FUNCTION_BLOCK basicUCT (* Logica unica da UCT Fast (Modbus TCP) e da bomba de gordura com a valvula de lavagem *)
  (* Standard: 61499-2 *)
  (* Version 1.7, 04/11/2026, Hidryco, Hidryco, 1.7: stsLigado para a IO List da Nereda. 1.6: nivel da peneira e velocidades da UCT em % direto (0-100); o 0-16000 da tabela e so o limite do registrador. IHM em Hz (60 Hz = 100 %). 1.5: velocidades dos equipamentos da UCT e da bomba de gordura em Hz (16000 = 60 Hz); conversao no CLP. 1.4: CNF_HMI tambem sai quando muda so a palavra de disponibilidade (STS_HABILITADA). 1.0: UCT Fast (memorial PR-809) por Modbus TCP - leitura de estado, comandos manuais e automaticos por evento, reset, disponibilidade para a EEE Bruto, bomba de gordura e valvula de lavagem *)
  PACKAGE Hidryco.HidrycoLib;
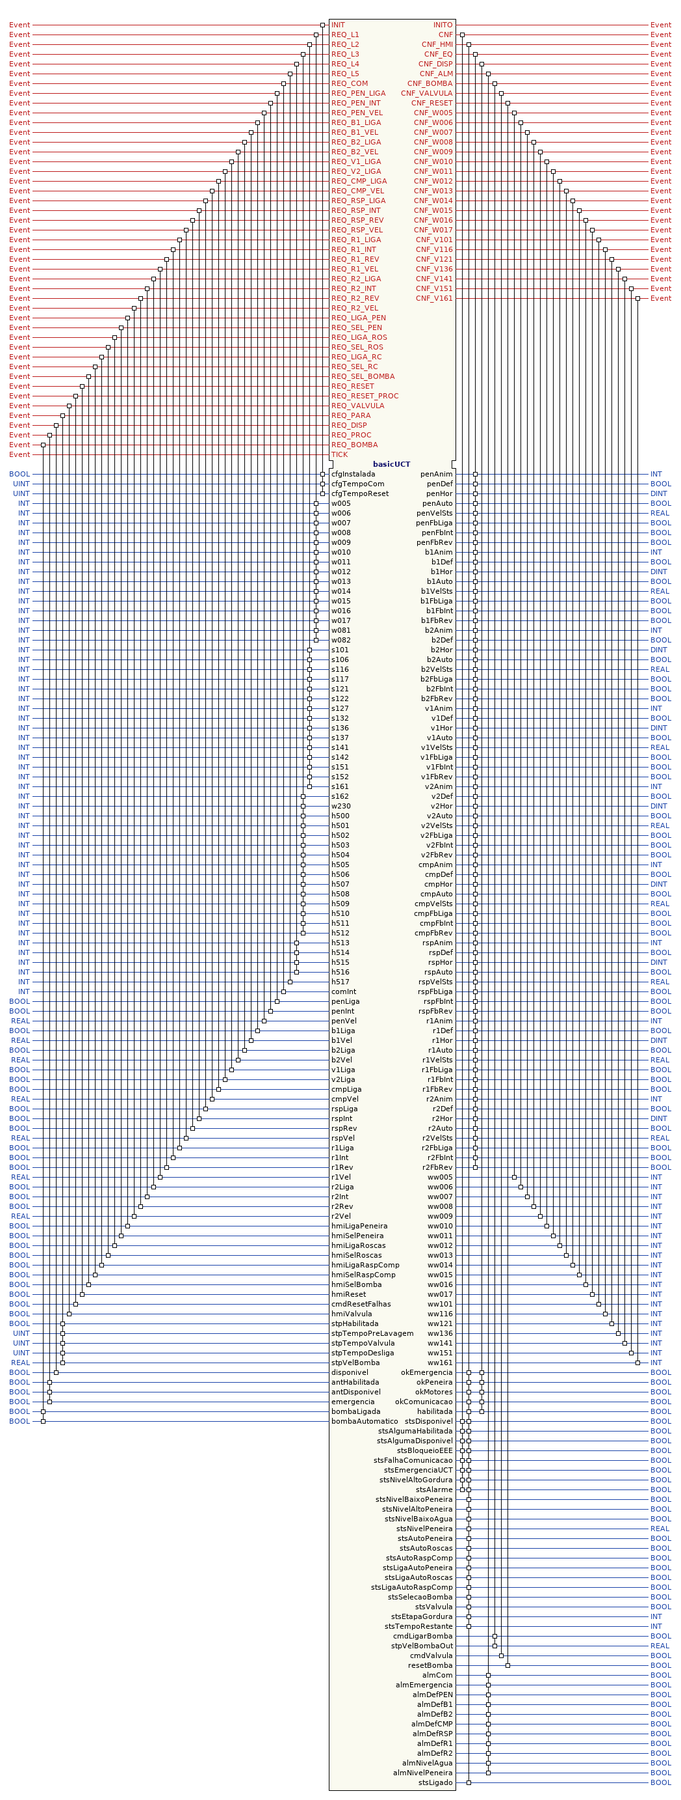
  EVENT_INPUT
    INIT WITH cfgInstalada, cfgTempoCom, cfgTempoReset; (* Inicializacao *)
    REQ_L1 WITH w005, w006, w007, w008, w009, w010, w011, w012, w013, w014, w015, w016, w017, w081, w082; (* Leitura Modbus (grupo 1) *)
    REQ_L2 WITH s101, s106, s116, s117, s121, s122, s127, s132, s136, s137, s141, s142, s151, s152, s161; (* Leitura Modbus (grupo 2) *)
    REQ_L3 WITH s162, w230, h500, h501, h502, h503, h504, h505, h506, h507, h508, h509, h510, h511, h512; (* Leitura Modbus (grupo 3) *)
    REQ_L4 WITH h513, h514, h515, h516; (* Leitura Modbus (grupo 4) *)
    REQ_L5 WITH h517; (* Leitura Modbus (grupo 5) *)
    REQ_COM WITH comInt; (* Comunicacao *)
    REQ_PEN_LIGA WITH penLiga; (* Peneira rotativa: liga manual *)
    REQ_PEN_INT WITH penInt; (* Peneira rotativa: intermitente *)
    REQ_PEN_VEL WITH penVel; (* Peneira rotativa: velocidade (%) *)
    REQ_B1_LIGA WITH b1Liga; (* Bomba 1 de higienização da peneira: liga manual *)
    REQ_B1_VEL WITH b1Vel; (* Bomba 1 de higienização da peneira: velocidade (%) *)
    REQ_B2_LIGA WITH b2Liga; (* Bomba 2 de higienização da peneira: liga manual *)
    REQ_B2_VEL WITH b2Vel; (* Bomba 2 de higienização da peneira: velocidade (%) *)
    REQ_V1_LIGA WITH v1Liga; (* Válvula 1 - higienização do cesto da peneira: liga manual *)
    REQ_V2_LIGA WITH v2Liga; (* Válvula 2 - higienização da rosca da peneira: liga manual *)
    REQ_CMP_LIGA WITH cmpLiga; (* Compressor de ar: liga manual *)
    REQ_CMP_VEL WITH cmpVel; (* Compressor de ar: velocidade (%) *)
    REQ_RSP_LIGA WITH rspLiga; (* Raspador de gordura: liga manual *)
    REQ_RSP_INT WITH rspInt; (* Raspador de gordura: intermitente *)
    REQ_RSP_REV WITH rspRev; (* Raspador de gordura: reversao *)
    REQ_RSP_VEL WITH rspVel; (* Raspador de gordura: velocidade (%) *)
    REQ_R1_LIGA WITH r1Liga; (* Rosca 1 - horizontal: liga manual *)
    REQ_R1_INT WITH r1Int; (* Rosca 1 - horizontal: intermitente *)
    REQ_R1_REV WITH r1Rev; (* Rosca 1 - horizontal: reversao *)
    REQ_R1_VEL WITH r1Vel; (* Rosca 1 - horizontal: velocidade (%) *)
    REQ_R2_LIGA WITH r2Liga; (* Rosca 2 - inclinada: liga manual *)
    REQ_R2_INT WITH r2Int; (* Rosca 2 - inclinada: intermitente *)
    REQ_R2_REV WITH r2Rev; (* Rosca 2 - inclinada: reversao *)
    REQ_R2_VEL WITH r2Vel; (* Rosca 2 - inclinada: velocidade (%) *)
    REQ_LIGA_PEN WITH hmiLigaPeneira; (* cmdLigaSubsistemaPeneira *)
    REQ_SEL_PEN WITH hmiSelPeneira; (* cmdSelecaoSubsistemaPeneira *)
    REQ_LIGA_ROS WITH hmiLigaRoscas; (* cmdLigaSubsistemaRoscas *)
    REQ_SEL_ROS WITH hmiSelRoscas; (* cmdSelecaoSubsistemaRoscas *)
    REQ_LIGA_RC WITH hmiLigaRaspComp; (* cmdLigaSubsistemaRaspComp *)
    REQ_SEL_RC WITH hmiSelRaspComp; (* cmdSelecaoSubsistemaRaspComp *)
    REQ_SEL_BOMBA WITH hmiSelBomba; (* cmdSelecaoBombaHigienizacao *)
    REQ_RESET WITH hmiReset; (* Reset pela IHM *)
    REQ_RESET_PROC WITH cmdResetFalhas; (* Reset pelo processo *)
    REQ_VALVULA WITH hmiValvula; (* Valvula de lavagem manual *)
    REQ_PARA WITH stpHabilitada, stpTempoPreLavagem, stpTempoValvula, stpTempoDesliga, stpVelBomba; (* Parametros (persistentes) *)
    REQ_DISP WITH disponivel; (* Resultado do AND de disponibilidade *)
    REQ_PROC WITH antHabilitada, antDisponivel, emergencia; (* Cadeia das UCTs e emergencia *)
    REQ_BOMBA WITH bombaLigada, bombaAutomatico; (* Estado da bomba de gordura *)
    TICK; (* Base de tempo de 1 s (E_CYCLE) *)
  END_EVENT
  EVENT_OUTPUT
    INITO; (* Inicializacao concluida *)
    CNF WITH stsDisponivel, stsAlgumaHabilitada, stsAlgumaDisponivel, stsBloqueioEEE, stsFalhaComunicacao, stsEmergenciaUCT, stsNivelAltoGordura, stsAlarme; (* Processo (na mudanca) *)
    CNF_HMI WITH stsDisponivel, stsAlgumaHabilitada, stsAlgumaDisponivel, stsBloqueioEEE, stsFalhaComunicacao, stsEmergenciaUCT, stsNivelAltoGordura, stsAlarme, stsNivelBaixoPeneira, stsNivelAltoPeneira, stsNivelBaixoAgua, stsNivelPeneira, stsAutoPeneira, stsAutoRoscas, stsAutoRaspComp, stsLigaAutoPeneira, stsLigaAutoRoscas, stsLigaAutoRaspComp, stsSelecaoBomba, stsValvula, stsEtapaGordura, stsTempoRestante, okEmergencia, okPeneira, okMotores, okComunicacao, habilitada, stsLigado; (* IHM da UCT (na mudanca) *)
    CNF_EQ WITH penAnim, penDef, penHor, penAuto, penVelSts, penFbLiga, penFbInt, penFbRev, b1Anim, b1Def, b1Hor, b1Auto, b1VelSts, b1FbLiga, b1FbInt, b1FbRev, b2Anim, b2Def, b2Hor, b2Auto, b2VelSts, b2FbLiga, b2FbInt, b2FbRev, v1Anim, v1Def, v1Hor, v1Auto, v1VelSts, v1FbLiga, v1FbInt, v1FbRev, v2Anim, v2Def, v2Hor, v2Auto, v2VelSts, v2FbLiga, v2FbInt, v2FbRev, cmpAnim, cmpDef, cmpHor, cmpAuto, cmpVelSts, cmpFbLiga, cmpFbInt, cmpFbRev, rspAnim, rspDef, rspHor, rspAuto, rspVelSts, rspFbLiga, rspFbInt, rspFbRev, r1Anim, r1Def, r1Hor, r1Auto, r1VelSts, r1FbLiga, r1FbInt, r1FbRev, r2Anim, r2Def, r2Hor, r2Auto, r2VelSts, r2FbLiga, r2FbInt, r2FbRev; (* IHM dos equipamentos (na mudanca) *)
    CNF_DISP WITH okEmergencia, okPeneira, okMotores, okComunicacao, habilitada; (* Condicoes para o AND de disponibilidade (na mudanca) *)
    CNF_ALM WITH almCom, almEmergencia, almDefPEN, almDefB1, almDefB2, almDefCMP, almDefRSP, almDefR1, almDefR2, almNivelAgua, almNivelPeneira; (* Alarmes para os ALARM_BIT (na mudanca) *)
    CNF_BOMBA WITH cmdLigarBomba, stpVelBombaOut; (* Bomba de gordura (na mudanca) *)
    CNF_VALVULA WITH cmdValvula; (* Valvula de lavagem (na mudanca) *)
    CNF_RESET WITH resetBomba; (* Reset da bomba de gordura *)
    CNF_W005 WITH ww005; (* Escreve 40005 na UCT *)
    CNF_W006 WITH ww006; (* Escreve 40006 na UCT *)
    CNF_W007 WITH ww007; (* Escreve 40007 na UCT *)
    CNF_W008 WITH ww008; (* Escreve 40008 na UCT *)
    CNF_W009 WITH ww009; (* Escreve 40009 na UCT *)
    CNF_W010 WITH ww010; (* Escreve 40010 na UCT *)
    CNF_W011 WITH ww011; (* Escreve 40011 na UCT *)
    CNF_W012 WITH ww012; (* Escreve 40012 na UCT *)
    CNF_W013 WITH ww013; (* Escreve 40013 na UCT *)
    CNF_W014 WITH ww014; (* Escreve 40014 na UCT *)
    CNF_W015 WITH ww015; (* Escreve 40015 na UCT *)
    CNF_W016 WITH ww016; (* Escreve 40016 na UCT *)
    CNF_W017 WITH ww017; (* Escreve 40017 na UCT *)
    CNF_V101 WITH ww101; (* Escreve 40101 na UCT *)
    CNF_V116 WITH ww116; (* Escreve 40116 na UCT *)
    CNF_V121 WITH ww121; (* Escreve 40121 na UCT *)
    CNF_V136 WITH ww136; (* Escreve 40136 na UCT *)
    CNF_V141 WITH ww141; (* Escreve 40141 na UCT *)
    CNF_V151 WITH ww151; (* Escreve 40151 na UCT *)
    CNF_V161 WITH ww161; (* Escreve 40161 na UCT *)
  END_EVENT
  VAR_INPUT
    cfgInstalada : BOOL := TRUE; (* FALSE = UCT ainda nao existe em campo (sem comunicacao, sem alarmes, fora do bloqueio da EEE) *)
    cfgTempoCom : UINT := 10; (* Tempo (s) sem comunicacao com a UCT para confirmar a falha *)
    cfgTempoReset : UINT := 2; (* Tempo (s) do pulso de reset escrito na UCT (40005.3) *)
    w005 : INT; (* Modbus UCT 40005 *)
    w006 : INT; (* Modbus UCT 40006 *)
    w007 : INT; (* Modbus UCT 40007 *)
    w008 : INT; (* Modbus UCT 40008 *)
    w009 : INT; (* Modbus UCT 40009 *)
    w010 : INT; (* Modbus UCT 40010 *)
    w011 : INT; (* Modbus UCT 40011 *)
    w012 : INT; (* Modbus UCT 40012 *)
    w013 : INT; (* Modbus UCT 40013 *)
    w014 : INT; (* Modbus UCT 40014 *)
    w015 : INT; (* Modbus UCT 40015 *)
    w016 : INT; (* Modbus UCT 40016 *)
    w017 : INT; (* Modbus UCT 40017 *)
    w081 : INT; (* Modbus UCT 40081 *)
    w082 : INT; (* Modbus UCT 40082 *)
    s101 : INT; (* Modbus UCT 40101 *)
    s106 : INT; (* Modbus UCT 40106 *)
    s116 : INT; (* Modbus UCT 40116 *)
    s117 : INT; (* Modbus UCT 40117 *)
    s121 : INT; (* Modbus UCT 40121 *)
    s122 : INT; (* Modbus UCT 40122 *)
    s127 : INT; (* Modbus UCT 40127 *)
    s132 : INT; (* Modbus UCT 40132 *)
    s136 : INT; (* Modbus UCT 40136 *)
    s137 : INT; (* Modbus UCT 40137 *)
    s141 : INT; (* Modbus UCT 40141 *)
    s142 : INT; (* Modbus UCT 40142 *)
    s151 : INT; (* Modbus UCT 40151 *)
    s152 : INT; (* Modbus UCT 40152 *)
    s161 : INT; (* Modbus UCT 40161 *)
    s162 : INT; (* Modbus UCT 40162 *)
    w230 : INT; (* Modbus UCT 40230 *)
    h500 : INT; (* Modbus UCT 40500 *)
    h501 : INT; (* Modbus UCT 40501 *)
    h502 : INT; (* Modbus UCT 40502 *)
    h503 : INT; (* Modbus UCT 40503 *)
    h504 : INT; (* Modbus UCT 40504 *)
    h505 : INT; (* Modbus UCT 40505 *)
    h506 : INT; (* Modbus UCT 40506 *)
    h507 : INT; (* Modbus UCT 40507 *)
    h508 : INT; (* Modbus UCT 40508 *)
    h509 : INT; (* Modbus UCT 40509 *)
    h510 : INT; (* Modbus UCT 40510 *)
    h511 : INT; (* Modbus UCT 40511 *)
    h512 : INT; (* Modbus UCT 40512 *)
    h513 : INT; (* Modbus UCT 40513 *)
    h514 : INT; (* Modbus UCT 40514 *)
    h515 : INT; (* Modbus UCT 40515 *)
    h516 : INT; (* Modbus UCT 40516 *)
    h517 : INT; (* Modbus UCT 40517 *)
    comInt : INT; (* connStatusInt do escravo Modbus da UCT (1 = online) *)
    penLiga : BOOL; (* IHM: Peneira rotativa: liga manual *)
    penInt : BOOL; (* IHM: Peneira rotativa: intermitente *)
    penVel : REAL; (* IHM: Peneira rotativa: velocidade (%) *)
    b1Liga : BOOL; (* IHM: Bomba 1 de higienização da peneira: liga manual *)
    b1Vel : REAL; (* IHM: Bomba 1 de higienização da peneira: velocidade (%) *)
    b2Liga : BOOL; (* IHM: Bomba 2 de higienização da peneira: liga manual *)
    b2Vel : REAL; (* IHM: Bomba 2 de higienização da peneira: velocidade (%) *)
    v1Liga : BOOL; (* IHM: Válvula 1 - higienização do cesto da peneira: liga manual *)
    v2Liga : BOOL; (* IHM: Válvula 2 - higienização da rosca da peneira: liga manual *)
    cmpLiga : BOOL; (* IHM: Compressor de ar: liga manual *)
    cmpVel : REAL; (* IHM: Compressor de ar: velocidade (%) *)
    rspLiga : BOOL; (* IHM: Raspador de gordura: liga manual *)
    rspInt : BOOL; (* IHM: Raspador de gordura: intermitente *)
    rspRev : BOOL; (* IHM: Raspador de gordura: reversao *)
    rspVel : REAL; (* IHM: Raspador de gordura: velocidade (%) *)
    r1Liga : BOOL; (* IHM: Rosca 1 - horizontal: liga manual *)
    r1Int : BOOL; (* IHM: Rosca 1 - horizontal: intermitente *)
    r1Rev : BOOL; (* IHM: Rosca 1 - horizontal: reversao *)
    r1Vel : REAL; (* IHM: Rosca 1 - horizontal: velocidade (%) *)
    r2Liga : BOOL; (* IHM: Rosca 2 - inclinada: liga manual *)
    r2Int : BOOL; (* IHM: Rosca 2 - inclinada: intermitente *)
    r2Rev : BOOL; (* IHM: Rosca 2 - inclinada: reversao *)
    r2Vel : REAL; (* IHM: Rosca 2 - inclinada: velocidade (%) *)
    hmiLigaPeneira : BOOL; (* IHM: cmdLigaSubsistemaPeneira *)
    hmiSelPeneira : BOOL; (* IHM: cmdSelecaoSubsistemaPeneira *)
    hmiLigaRoscas : BOOL; (* IHM: cmdLigaSubsistemaRoscas *)
    hmiSelRoscas : BOOL; (* IHM: cmdSelecaoSubsistemaRoscas *)
    hmiLigaRaspComp : BOOL; (* IHM: cmdLigaSubsistemaRaspComp *)
    hmiSelRaspComp : BOOL; (* IHM: cmdSelecaoSubsistemaRaspComp *)
    hmiSelBomba : BOOL; (* IHM: cmdSelecaoBombaHigienizacao *)
    hmiReset : BOOL; (* IHM: reset (reconhece e reseta a UCT e a bomba de gordura) *)
    cmdResetFalhas : BOOL; (* Processo: reset (com E_RESET_FALHAS) *)
    hmiValvula : BOOL; (* IHM: valvula de lavagem aberta (TRUE) / fechada (FALSE) - so com a bomba de gordura fora do automatico *)
    stpHabilitada : BOOL; (* IHM (persistente): UCT habilitada no bloqueio da EEE Bruto (desabilitada nao conta) *)
    stpTempoPreLavagem : UINT; (* IHM (persistente): Tempo (s) com a valvula de lavagem aberta antes de ligar a bomba de gordura (0 = liga junto) *)
    stpTempoValvula : UINT; (* IHM (persistente): Tempo (s) que a valvula fica aberta depois que a bomba liga (0 = fecha na partida) *)
    stpTempoDesliga : UINT; (* IHM (persistente): Tempo (s) que a bomba de gordura continua ligada depois que o nivel alto do tanque abaixa *)
    stpVelBomba : REAL; (* IHM (persistente): Velocidade da bomba de gordura em automatico (%) *)
    disponivel : BOOL; (* Saida do bloco AND editavel: UCT disponivel *)
    antHabilitada : BOOL; (* UCT anterior na cadeia: alguma UCT habilitada *)
    antDisponivel : BOOL; (* UCT anterior na cadeia: alguma UCT disponivel *)
    emergencia : BOOL; (* Emergencia pelo processo (fecha a valvula de lavagem) *)
    bombaLigada : BOOL; (* Bomba de gordura ligada (Motor_Generico.stsLigado) *)
    bombaAutomatico : BOOL; (* Bomba de gordura em automatico (Motor_Generico.stsAutomatico) *)
  END_VAR
  VAR_OUTPUT
    penAnim : INT; (* Peneira rotativa: 0 desligado, 1 ligado, 2 falha, 3 manutencao, 4 sem comunicacao *)
    penDef : BOOL; (* Peneira rotativa: defeito *)
    penHor : DINT; (* Peneira rotativa: horimetro (h) *)
    penAuto : BOOL; (* Peneira rotativa: subsistema em automatico *)
    penVelSts : REAL; (* Peneira rotativa: velocidade (%) *)
    penFbLiga : BOOL; (* Peneira rotativa: liga em vigor *)
    penFbInt : BOOL; (* Peneira rotativa: intermitente em vigor *)
    penFbRev : BOOL; (* Peneira rotativa: reversao em vigor *)
    b1Anim : INT; (* Bomba 1 de higienização da peneira: 0 desligado, 1 ligado, 2 falha, 3 manutencao, 4 sem comunicacao *)
    b1Def : BOOL; (* Bomba 1 de higienização da peneira: defeito *)
    b1Hor : DINT; (* Bomba 1 de higienização da peneira: horimetro (h) *)
    b1Auto : BOOL; (* Bomba 1 de higienização da peneira: subsistema em automatico *)
    b1VelSts : REAL; (* Bomba 1 de higienização da peneira: velocidade (%) *)
    b1FbLiga : BOOL; (* Bomba 1 de higienização da peneira: liga em vigor *)
    b1FbInt : BOOL; (* Bomba 1 de higienização da peneira: intermitente em vigor *)
    b1FbRev : BOOL; (* Bomba 1 de higienização da peneira: reversao em vigor *)
    b2Anim : INT; (* Bomba 2 de higienização da peneira: 0 desligado, 1 ligado, 2 falha, 3 manutencao, 4 sem comunicacao *)
    b2Def : BOOL; (* Bomba 2 de higienização da peneira: defeito *)
    b2Hor : DINT; (* Bomba 2 de higienização da peneira: horimetro (h) *)
    b2Auto : BOOL; (* Bomba 2 de higienização da peneira: subsistema em automatico *)
    b2VelSts : REAL; (* Bomba 2 de higienização da peneira: velocidade (%) *)
    b2FbLiga : BOOL; (* Bomba 2 de higienização da peneira: liga em vigor *)
    b2FbInt : BOOL; (* Bomba 2 de higienização da peneira: intermitente em vigor *)
    b2FbRev : BOOL; (* Bomba 2 de higienização da peneira: reversao em vigor *)
    v1Anim : INT; (* Válvula 1 - higienização do cesto da peneira: 0 desligado, 1 ligado, 2 falha, 3 manutencao, 4 sem comunicacao *)
    v1Def : BOOL; (* Válvula 1 - higienização do cesto da peneira: defeito *)
    v1Hor : DINT; (* Válvula 1 - higienização do cesto da peneira: horimetro (h) *)
    v1Auto : BOOL; (* Válvula 1 - higienização do cesto da peneira: subsistema em automatico *)
    v1VelSts : REAL; (* Válvula 1 - higienização do cesto da peneira: velocidade (%) *)
    v1FbLiga : BOOL; (* Válvula 1 - higienização do cesto da peneira: liga em vigor *)
    v1FbInt : BOOL; (* Válvula 1 - higienização do cesto da peneira: intermitente em vigor *)
    v1FbRev : BOOL; (* Válvula 1 - higienização do cesto da peneira: reversao em vigor *)
    v2Anim : INT; (* Válvula 2 - higienização da rosca da peneira: 0 desligado, 1 ligado, 2 falha, 3 manutencao, 4 sem comunicacao *)
    v2Def : BOOL; (* Válvula 2 - higienização da rosca da peneira: defeito *)
    v2Hor : DINT; (* Válvula 2 - higienização da rosca da peneira: horimetro (h) *)
    v2Auto : BOOL; (* Válvula 2 - higienização da rosca da peneira: subsistema em automatico *)
    v2VelSts : REAL; (* Válvula 2 - higienização da rosca da peneira: velocidade (%) *)
    v2FbLiga : BOOL; (* Válvula 2 - higienização da rosca da peneira: liga em vigor *)
    v2FbInt : BOOL; (* Válvula 2 - higienização da rosca da peneira: intermitente em vigor *)
    v2FbRev : BOOL; (* Válvula 2 - higienização da rosca da peneira: reversao em vigor *)
    cmpAnim : INT; (* Compressor de ar: 0 desligado, 1 ligado, 2 falha, 3 manutencao, 4 sem comunicacao *)
    cmpDef : BOOL; (* Compressor de ar: defeito *)
    cmpHor : DINT; (* Compressor de ar: horimetro (h) *)
    cmpAuto : BOOL; (* Compressor de ar: subsistema em automatico *)
    cmpVelSts : REAL; (* Compressor de ar: velocidade (%) *)
    cmpFbLiga : BOOL; (* Compressor de ar: liga em vigor *)
    cmpFbInt : BOOL; (* Compressor de ar: intermitente em vigor *)
    cmpFbRev : BOOL; (* Compressor de ar: reversao em vigor *)
    rspAnim : INT; (* Raspador de gordura: 0 desligado, 1 ligado, 2 falha, 3 manutencao, 4 sem comunicacao *)
    rspDef : BOOL; (* Raspador de gordura: defeito *)
    rspHor : DINT; (* Raspador de gordura: horimetro (h) *)
    rspAuto : BOOL; (* Raspador de gordura: subsistema em automatico *)
    rspVelSts : REAL; (* Raspador de gordura: velocidade (%) *)
    rspFbLiga : BOOL; (* Raspador de gordura: liga em vigor *)
    rspFbInt : BOOL; (* Raspador de gordura: intermitente em vigor *)
    rspFbRev : BOOL; (* Raspador de gordura: reversao em vigor *)
    r1Anim : INT; (* Rosca 1 - horizontal: 0 desligado, 1 ligado, 2 falha, 3 manutencao, 4 sem comunicacao *)
    r1Def : BOOL; (* Rosca 1 - horizontal: defeito *)
    r1Hor : DINT; (* Rosca 1 - horizontal: horimetro (h) *)
    r1Auto : BOOL; (* Rosca 1 - horizontal: subsistema em automatico *)
    r1VelSts : REAL; (* Rosca 1 - horizontal: velocidade (%) *)
    r1FbLiga : BOOL; (* Rosca 1 - horizontal: liga em vigor *)
    r1FbInt : BOOL; (* Rosca 1 - horizontal: intermitente em vigor *)
    r1FbRev : BOOL; (* Rosca 1 - horizontal: reversao em vigor *)
    r2Anim : INT; (* Rosca 2 - inclinada: 0 desligado, 1 ligado, 2 falha, 3 manutencao, 4 sem comunicacao *)
    r2Def : BOOL; (* Rosca 2 - inclinada: defeito *)
    r2Hor : DINT; (* Rosca 2 - inclinada: horimetro (h) *)
    r2Auto : BOOL; (* Rosca 2 - inclinada: subsistema em automatico *)
    r2VelSts : REAL; (* Rosca 2 - inclinada: velocidade (%) *)
    r2FbLiga : BOOL; (* Rosca 2 - inclinada: liga em vigor *)
    r2FbInt : BOOL; (* Rosca 2 - inclinada: intermitente em vigor *)
    r2FbRev : BOOL; (* Rosca 2 - inclinada: reversao em vigor *)
    ww005 : INT; (* Palavra escrita na UCT: 40005 *)
    ww006 : INT; (* Palavra escrita na UCT: 40006 *)
    ww007 : INT; (* Palavra escrita na UCT: 40007 *)
    ww008 : INT; (* Palavra escrita na UCT: 40008 *)
    ww009 : INT; (* Palavra escrita na UCT: 40009 *)
    ww010 : INT; (* Palavra escrita na UCT: 40010 *)
    ww011 : INT; (* Palavra escrita na UCT: 40011 *)
    ww012 : INT; (* Palavra escrita na UCT: 40012 *)
    ww013 : INT; (* Palavra escrita na UCT: 40013 *)
    ww014 : INT; (* Palavra escrita na UCT: 40014 *)
    ww015 : INT; (* Palavra escrita na UCT: 40015 *)
    ww016 : INT; (* Palavra escrita na UCT: 40016 *)
    ww017 : INT; (* Palavra escrita na UCT: 40017 *)
    ww101 : INT; (* Palavra escrita na UCT: 40101 *)
    ww116 : INT; (* Palavra escrita na UCT: 40116 *)
    ww121 : INT; (* Palavra escrita na UCT: 40121 *)
    ww136 : INT; (* Palavra escrita na UCT: 40136 *)
    ww141 : INT; (* Palavra escrita na UCT: 40141 *)
    ww151 : INT; (* Palavra escrita na UCT: 40151 *)
    ww161 : INT; (* Palavra escrita na UCT: 40161 *)
    okEmergencia : BOOL; (* UCT sem emergencia *)
    okPeneira : BOOL; (* Peneira sem defeito *)
    okMotores : BOOL; (* Bombas de higienizacao, roscas, raspador e compressor sem defeito *)
    okComunicacao : BOOL; (* Comunicacao com a UCT ok *)
    habilitada : BOOL; (* UCT instalada e habilitada *)
    stsDisponivel : BOOL; (* UCT disponivel (saida do AND) *)
    stsAlgumaHabilitada : BOOL; (* Esta UCT ou alguma anterior habilitada *)
    stsAlgumaDisponivel : BOOL; (* Esta UCT ou alguma anterior disponivel *)
    stsBloqueioEEE : BOOL; (* Bloqueio do automatico da EEE Bruto: ha UCT habilitada e nenhuma disponivel *)
    stsFalhaComunicacao : BOOL; (* Falha de comunicacao com a UCT *)
    stsEmergenciaUCT : BOOL; (* Emergencia acionada na UCT *)
    stsNivelAltoGordura : BOOL; (* Nivel alto do tanque de gordura (UCT) *)
    stsAlarme : BOOL; (* Algum alarme da UCT *)
    stsNivelBaixoPeneira : BOOL; (* Nivel baixo da peneira *)
    stsNivelAltoPeneira : BOOL; (* Nivel alto da peneira *)
    stsNivelBaixoAgua : BOOL; (* Nivel baixo do tanque de agua *)
    stsNivelPeneira : REAL; (* Nivel da peneira (%) *)
    stsAutoPeneira : BOOL; (* Subsistema peneira e higienização em automatico *)
    stsAutoRoscas : BOOL; (* Subsistema roscas em automatico *)
    stsAutoRaspComp : BOOL; (* Subsistema raspador e compressor em automatico *)
    stsLigaAutoPeneira : BOOL; (* Subsistema peneira e higienização: liga automatico em vigor *)
    stsLigaAutoRoscas : BOOL; (* Subsistema roscas: liga automatico em vigor *)
    stsLigaAutoRaspComp : BOOL; (* Subsistema raspador e compressor: liga automatico em vigor *)
    stsSelecaoBomba : BOOL; (* Bomba de higienizacao selecionada: FALSE = bomba 1, TRUE = bomba 2 *)
    stsValvula : BOOL; (* Valvula de lavagem do tanque de gordura aberta *)
    stsEtapaGordura : INT; (* Bomba de gordura: 0 parada, 1 pre-lavagem, 2 bombeando, 3 nivel normal - contando para desligar, 4 fora do automatico *)
    stsTempoRestante : INT; (* Tempo restante (s) da etapa da bomba de gordura *)
    cmdLigarBomba : BOOL; (* Bomba de gordura: liga em automatico (Motor_Generico.cmdLigarAutomatico) *)
    stpVelBombaOut : REAL; (* Bomba de gordura: velocidade em automatico (%) *)
    cmdValvula : BOOL; (* Valvula de lavagem: saida digital (symlink ${PATH}cmdValvulaLavagem) *)
    resetBomba : BOOL; (* Reset da bomba de gordura (com CNF_RESET) *)
    almCom : BOOL; (* ALARM_BIT Falha de comunicação com a UCT *)
    almEmergencia : BOOL; (* ALARM_BIT Emergência acionada na UCT *)
    almDefPEN : BOOL; (* ALARM_BIT Defeito: Peneira rotativa *)
    almDefB1 : BOOL; (* ALARM_BIT Defeito: Bomba 1 de higienização da peneira *)
    almDefB2 : BOOL; (* ALARM_BIT Defeito: Bomba 2 de higienização da peneira *)
    almDefCMP : BOOL; (* ALARM_BIT Defeito: Compressor de ar *)
    almDefRSP : BOOL; (* ALARM_BIT Defeito: Raspador de gordura *)
    almDefR1 : BOOL; (* ALARM_BIT Defeito: Rosca 1 - horizontal *)
    almDefR2 : BOOL; (* ALARM_BIT Defeito: Rosca 2 - inclinada *)
    almNivelAgua : BOOL; (* ALARM_BIT Nível baixo do tanque de água de higienização da UCT *)
    almNivelPeneira : BOOL; (* ALARM_BIT Nível alto na peneira da UCT *)
    stsLigado : BOOL; (* Algum subsistema com liga-automatico (peneira, roscas ou raspador/compressor) *)
  END_VAR
  VAR
    initDone : BOOL;
    initPass : BOOL;
    bComRecebida : BOOL; (* Ja houve leitura do connStatusInt *)
    bLeitura : BOOL; (* Ja houve leitura das palavras de comando *)
    bComOK : BOOL; (* Comunicando agora *)
    uSegCom : UDINT;
    uSegReset : UINT; (* Segundos do pulso de reset *)
    bReset : BOOL;
    w81 : WORD;
    w82 : WORD;
    bNivelAltoG : BOOL; (* Nivel alto do tanque de gordura valido *)
    uEtapa : INT; (* Etapa da bomba de gordura *)
    uSegEtapa : UDINT; (* Segundos na etapa *)
    uSegValv : UDINT; (* Segundos com a bomba ligada *)
    bValvAuto : BOOL; (* Valvula pedida pela sequencia *)
    bMudou : BOOL;
    wD : WORD;
    oldD : WORD := 16#FFFF;
    wP : DWORD;
    oldP : DWORD := 16#FFFFFFFF;
    wA : WORD;
    oldA : WORD := 16#FFFF;
    oldLigB : BOOL;
    oldVelB : REAL := -1.0;
    oldValv : BOOL;
    img005 : WORD; (* Imagem da palavra 40005 (lida da UCT, alterada so no bit comandado) *)
    img006 : WORD; (* Imagem da palavra 40006 (lida da UCT, alterada so no bit comandado) *)
    img007 : WORD; (* Imagem da palavra 40007 (lida da UCT, alterada so no bit comandado) *)
    img008 : WORD; (* Imagem da palavra 40008 (lida da UCT, alterada so no bit comandado) *)
    img009 : WORD; (* Imagem da palavra 40009 (lida da UCT, alterada so no bit comandado) *)
    img010 : WORD; (* Imagem da palavra 40010 (lida da UCT, alterada so no bit comandado) *)
    img011 : WORD; (* Imagem da palavra 40011 (lida da UCT, alterada so no bit comandado) *)
    img012 : WORD; (* Imagem da palavra 40012 (lida da UCT, alterada so no bit comandado) *)
    img013 : WORD; (* Imagem da palavra 40013 (lida da UCT, alterada so no bit comandado) *)
    img014 : WORD; (* Imagem da palavra 40014 (lida da UCT, alterada so no bit comandado) *)
    img015 : WORD; (* Imagem da palavra 40015 (lida da UCT, alterada so no bit comandado) *)
    img016 : WORD; (* Imagem da palavra 40016 (lida da UCT, alterada so no bit comandado) *)
    img017 : WORD; (* Imagem da palavra 40017 (lida da UCT, alterada so no bit comandado) *)
    o_stsNivelPeneira : REAL := -1.0;
    o_stsEtapaGordura : INT := -1;
    o_stsTempoRestante : INT := -1;
    o_penAnim : INT := -1;
    o_penHor : DINT := -1;
    o_penVelSts : REAL := -1.0;
    o_b1Anim : INT := -1;
    o_b1Hor : DINT := -1;
    o_b1VelSts : REAL := -1.0;
    o_b2Anim : INT := -1;
    o_b2Hor : DINT := -1;
    o_b2VelSts : REAL := -1.0;
    o_v1Anim : INT := -1;
    o_v1Hor : DINT := -1;
    o_v1VelSts : REAL := -1.0;
    o_v2Anim : INT := -1;
    o_v2Hor : DINT := -1;
    o_v2VelSts : REAL := -1.0;
    o_cmpAnim : INT := -1;
    o_cmpHor : DINT := -1;
    o_cmpVelSts : REAL := -1.0;
    o_rspAnim : INT := -1;
    o_rspHor : DINT := -1;
    o_rspVelSts : REAL := -1.0;
    o_r1Anim : INT := -1;
    o_r1Hor : DINT := -1;
    o_r1VelSts : REAL := -1.0;
    o_r2Anim : INT := -1;
    o_r2Hor : DINT := -1;
    o_r2VelSts : REAL := -1.0;
    o_penDef : BOOL;
    o_penAuto : BOOL;
    o_penFbLiga : BOOL;
    o_penFbInt : BOOL;
    o_penFbRev : BOOL;
    o_b1Def : BOOL;
    o_b1Auto : BOOL;
    o_b1FbLiga : BOOL;
    o_b1FbInt : BOOL;
    o_b1FbRev : BOOL;
    o_b2Def : BOOL;
    o_b2Auto : BOOL;
    o_b2FbLiga : BOOL;
    o_b2FbInt : BOOL;
    o_b2FbRev : BOOL;
    o_v1Def : BOOL;
    o_v1Auto : BOOL;
    o_v1FbLiga : BOOL;
    o_v1FbInt : BOOL;
    o_v1FbRev : BOOL;
    o_v2Def : BOOL;
    o_v2Auto : BOOL;
    o_v2FbLiga : BOOL;
    o_v2FbInt : BOOL;
    o_v2FbRev : BOOL;
    o_cmpDef : BOOL;
    o_cmpAuto : BOOL;
    o_cmpFbLiga : BOOL;
    o_cmpFbInt : BOOL;
    o_cmpFbRev : BOOL;
    o_rspDef : BOOL;
    o_rspAuto : BOOL;
    o_rspFbLiga : BOOL;
    o_rspFbInt : BOOL;
    o_rspFbRev : BOOL;
    o_r1Def : BOOL;
    o_r1Auto : BOOL;
    o_r1FbLiga : BOOL;
    o_r1FbInt : BOOL;
    o_r1FbRev : BOOL;
    o_r2Def : BOOL;
    o_r2Auto : BOOL;
    o_r2FbLiga : BOOL;
    o_r2FbInt : BOOL;
    o_r2FbRev : BOOL;
  END_VAR
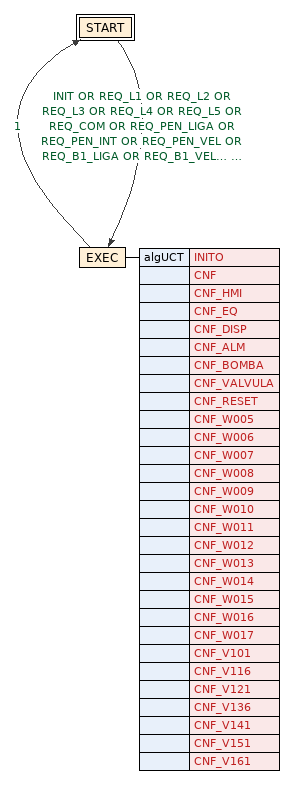
  EC_STATES
    START; (* Estado inicial *)
    EXEC : algUCT -> INITO, -> CNF, -> CNF_HMI, -> CNF_EQ, -> CNF_DISP, -> CNF_ALM, -> CNF_BOMBA, -> CNF_VALVULA, -> CNF_RESET, -> CNF_W005, -> CNF_W006, -> CNF_W007, -> CNF_W008, -> CNF_W009, -> CNF_W010, -> CNF_W011, -> CNF_W012, -> CNF_W013, -> CNF_W014, -> CNF_W015, -> CNF_W016, -> CNF_W017, -> CNF_V101, -> CNF_V116, -> CNF_V121, -> CNF_V136, -> CNF_V141, -> CNF_V151, -> CNF_V161; (* Executa a logica; o algoritmo decide quais eventos saem *)
  END_STATES
  EC_TRANSITIONS
    START TO EXEC := INIT OR REQ_L1 OR REQ_L2 OR REQ_L3 OR REQ_L4 OR REQ_L5 OR REQ_COM OR REQ_PEN_LIGA OR REQ_PEN_INT OR REQ_PEN_VEL OR REQ_B1_LIGA OR REQ_B1_VEL OR REQ_B2_LIGA OR REQ_B2_VEL OR REQ_V1_LIGA OR REQ_V2_LIGA OR REQ_CMP_LIGA OR REQ_CMP_VEL OR REQ_RSP_LIGA OR REQ_RSP_INT OR REQ_RSP_REV OR REQ_RSP_VEL OR REQ_R1_LIGA OR REQ_R1_INT OR REQ_R1_REV OR REQ_R1_VEL OR REQ_R2_LIGA OR REQ_R2_INT OR REQ_R2_REV OR REQ_R2_VEL OR REQ_LIGA_PEN OR REQ_SEL_PEN OR REQ_LIGA_ROS OR REQ_SEL_ROS OR REQ_LIGA_RC OR REQ_SEL_RC OR REQ_SEL_BOMBA OR REQ_RESET OR REQ_RESET_PROC OR REQ_VALVULA OR REQ_PARA OR REQ_DISP OR REQ_PROC OR REQ_BOMBA OR TICK;
    EXEC TO START := 1;
  END_TRANSITIONS
  ALGORITHM algUCT IN ST: (* Logica completa da UCT (um unico algoritmo) *)
(* =====================================================================
   basicUCT v1.0 - UCT Fast (tratamento preliminar) por Modbus TCP
   Padrao das bibliotecas Schneider: eventos de saida desligados no inicio e
   ligados so na mudanca; tempos pelo TICK de 1 s (E_CYCLE do CAT).
   - leitura: palavras de comando 40005..40017 (imagem), falhas 40081,
     niveis 40082, status/velocidade dos equipamentos 401xx, nivel da
     peneira 40230 (0-100 %, direto), horimetros 40500..40517 (DINT,
     palavra baixa no endereco menor);
   - escrita so quando o operador comanda (um evento por comando): o bit
     comandado e trocado na imagem lida e a palavra inteira e escrita
     (os outros bits ficam como a UCT informou); velocidade em Hz ->
     0-100 % (60 Hz = 100 %); reset = pulso de cfgTempoReset s em 40005.3;
   - disponibilidade: as condicoes vao para o bloco AND do CAT (editavel)
     e o resultado volta em "disponivel"; cadeia das UCTs: bloqueio da EEE
     Bruto so com UCT habilitada e nenhuma disponivel;
   - bomba de gordura (automatico): nivel alto do tanque de gordura ->
     abre a valvula de lavagem, espera stpTempoPreLavagem e liga a bomba;
     a valvula fecha stpTempoValvula s depois da partida; com o nivel
     normal conta stpTempoDesliga e desliga; fora do automatico a
     valvula segue o botao da IHM.
   ===================================================================== *)

(* ---- 0. Eventos de saida: so sai o que for ligado abaixo ---- *)
INITO := FALSE;
CNF := FALSE;
CNF_HMI := FALSE;
CNF_EQ := FALSE;
CNF_DISP := FALSE;
CNF_ALM := FALSE;
CNF_BOMBA := FALSE;
CNF_VALVULA := FALSE;
CNF_RESET := FALSE;
CNF_W005 := FALSE;
CNF_W006 := FALSE;
CNF_W007 := FALSE;
CNF_W008 := FALSE;
CNF_W009 := FALSE;
CNF_W010 := FALSE;
CNF_W011 := FALSE;
CNF_W012 := FALSE;
CNF_W013 := FALSE;
CNF_W014 := FALSE;
CNF_W015 := FALSE;
CNF_W016 := FALSE;
CNF_W017 := FALSE;
CNF_V101 := FALSE;
CNF_V116 := FALSE;
CNF_V121 := FALSE;
CNF_V136 := FALSE;
CNF_V141 := FALSE;
CNF_V151 := FALSE;
CNF_V161 := FALSE;

IF REQ_COM THEN
    bComRecebida := TRUE;
END_IF;
IF REQ_L1 THEN
    bLeitura := TRUE;
    img005 := INT_TO_WORD(w005);
    img006 := INT_TO_WORD(w006);
    img007 := INT_TO_WORD(w007);
    img008 := INT_TO_WORD(w008);
    img009 := INT_TO_WORD(w009);
    img010 := INT_TO_WORD(w010);
    img011 := INT_TO_WORD(w011);
    img012 := INT_TO_WORD(w012);
    img013 := INT_TO_WORD(w013);
    img014 := INT_TO_WORD(w014);
    img015 := INT_TO_WORD(w015);
    img016 := INT_TO_WORD(w016);
    img017 := INT_TO_WORD(w017);
END_IF;

(* ---- 1. Inicializacao ---- *)
IF INIT THEN
    initDone := TRUE;
    initPass := TRUE;
    INITO    := TRUE;
END_IF;
IF NOT initDone THEN
    RETURN;
END_IF;

(* ---- 2. Comunicacao (falha confirmada depois de cfgTempoCom s) ---- *)
bComOK := cfgInstalada AND bComRecebida AND comInt = 1;
IF cfgInstalada AND NOT bComOK THEN
    IF TICK AND uSegCom < UINT_TO_UDINT(cfgTempoCom) THEN
        uSegCom := uSegCom + 1;
    END_IF;
ELSE
    uSegCom := 0;
END_IF;
stsFalhaComunicacao := cfgInstalada AND NOT bComOK AND uSegCom >= UINT_TO_UDINT(cfgTempoCom);

(* ---- 3. Estado lido (com a comunicacao em falha os valores ficam congelados) ---- *)
w81 := INT_TO_WORD(w081);
w82 := INT_TO_WORD(w082);
stsEmergenciaUCT := bComOK AND ((w81 AND 16#0001) <> 16#0000);
stsNivelBaixoPeneira := bComOK AND ((w82 AND 16#0001) <> 16#0000);
stsNivelAltoPeneira := bComOK AND ((w82 AND 16#0002) <> 16#0000);
stsNivelBaixoAgua := bComOK AND ((w82 AND 16#0004) <> 16#0000);
stsNivelAltoGordura := bComOK AND ((w82 AND 16#0008) <> 16#0000);
stsNivelPeneira := INT_TO_REAL(w230);   (* % direto *)
stsAutoPeneira := (img015 AND 16#0004) <> 16#0000;
stsLigaAutoPeneira := (img015 AND 16#0001) <> 16#0000;
stsAutoRoscas := (img016 AND 16#0004) <> 16#0000;
stsLigaAutoRoscas := (img016 AND 16#0001) <> 16#0000;
stsAutoRaspComp := (img017 AND 16#0004) <> 16#0000;
stsLigaAutoRaspComp := (img017 AND 16#0001) <> 16#0000;
(* IO List da Nereda: UCT ligada = algum subsistema com liga-automatico *)
stsLigado := stsLigaAutoPeneira OR stsLigaAutoRoscas OR stsLigaAutoRaspComp;
stsSelecaoBomba := (img007 AND 16#0008) <> 16#0000;
(* Peneira rotativa *)
IF bComOK THEN
    penAnim := s106;
ELSE
    penAnim := 4;
END_IF;
penDef := bComOK AND ((w81 AND 16#0010) <> 16#0000);
penHor := DWORD_TO_DINT(SHL(WORD_TO_DWORD(INT_TO_WORD(h501)), 16) OR WORD_TO_DWORD(INT_TO_WORD(h500)));
penAuto := stsAutoPeneira;
penVelSts := INT_TO_REAL(s101) * 60.0 / 100.0;   (* Hz; UCT em % *)
penFbLiga := (img006 AND 16#0001) <> 16#0000;
penFbInt := (img006 AND 16#0020) <> 16#0000;
penFbRev := FALSE;
(* Bomba 1 de higienização da peneira *)
IF bComOK THEN
    b1Anim := s117;
ELSE
    b1Anim := 4;
END_IF;
b1Def := bComOK AND ((w81 AND 16#0004) <> 16#0000);
b1Hor := DWORD_TO_DINT(SHL(WORD_TO_DWORD(INT_TO_WORD(h503)), 16) OR WORD_TO_DWORD(INT_TO_WORD(h502)));
b1Auto := stsAutoPeneira;
b1VelSts := INT_TO_REAL(s116) * 60.0 / 100.0;   (* Hz; UCT em % *)
b1FbLiga := (img007 AND 16#0001) <> 16#0000;
b1FbInt := FALSE;
b1FbRev := FALSE;
(* Bomba 2 de higienização da peneira *)
IF bComOK THEN
    b2Anim := s122;
ELSE
    b2Anim := 4;
END_IF;
b2Def := bComOK AND ((w81 AND 16#0008) <> 16#0000);
b2Hor := DWORD_TO_DINT(SHL(WORD_TO_DWORD(INT_TO_WORD(h505)), 16) OR WORD_TO_DWORD(INT_TO_WORD(h504)));
b2Auto := stsAutoPeneira;
b2VelSts := INT_TO_REAL(s121) * 60.0 / 100.0;   (* Hz; UCT em % *)
b2FbLiga := (img008 AND 16#0001) <> 16#0000;
b2FbInt := FALSE;
b2FbRev := FALSE;
(* Válvula 1 - higienização do cesto da peneira *)
IF bComOK THEN
    v1Anim := s127;
ELSE
    v1Anim := 4;
END_IF;
v1Def := bComOK AND (s127 = 2);
v1Hor := DWORD_TO_DINT(SHL(WORD_TO_DWORD(INT_TO_WORD(h507)), 16) OR WORD_TO_DWORD(INT_TO_WORD(h506)));
v1Auto := stsAutoPeneira;
v1VelSts := 0.0;
v1FbLiga := (img009 AND 16#0001) <> 16#0000;
v1FbInt := FALSE;
v1FbRev := FALSE;
(* Válvula 2 - higienização da rosca da peneira *)
IF bComOK THEN
    v2Anim := s132;
ELSE
    v2Anim := 4;
END_IF;
v2Def := bComOK AND (s132 = 2);
v2Hor := DWORD_TO_DINT(SHL(WORD_TO_DWORD(INT_TO_WORD(h509)), 16) OR WORD_TO_DWORD(INT_TO_WORD(h508)));
v2Auto := stsAutoPeneira;
v2VelSts := 0.0;
v2FbLiga := (img010 AND 16#0001) <> 16#0000;
v2FbInt := FALSE;
v2FbRev := FALSE;
(* Compressor de ar *)
IF bComOK THEN
    cmpAnim := s137;
ELSE
    cmpAnim := 4;
END_IF;
cmpDef := bComOK AND ((w81 AND 16#0100) <> 16#0000);
cmpHor := DWORD_TO_DINT(SHL(WORD_TO_DWORD(INT_TO_WORD(h511)), 16) OR WORD_TO_DWORD(INT_TO_WORD(h510)));
cmpAuto := stsAutoRaspComp;
cmpVelSts := INT_TO_REAL(s136) * 60.0 / 100.0;   (* Hz; UCT em % *)
cmpFbLiga := (img011 AND 16#0001) <> 16#0000;
cmpFbInt := FALSE;
cmpFbRev := FALSE;
(* Raspador de gordura *)
IF bComOK THEN
    rspAnim := s142;
ELSE
    rspAnim := 4;
END_IF;
rspDef := bComOK AND ((w81 AND 16#0080) <> 16#0000);
rspHor := DWORD_TO_DINT(SHL(WORD_TO_DWORD(INT_TO_WORD(h513)), 16) OR WORD_TO_DWORD(INT_TO_WORD(h512)));
rspAuto := stsAutoRaspComp;
rspVelSts := INT_TO_REAL(s141) * 60.0 / 100.0;   (* Hz; UCT em % *)
rspFbLiga := (img012 AND 16#0001) <> 16#0000;
rspFbInt := (img012 AND 16#0020) <> 16#0000;
rspFbRev := (img012 AND 16#0008) <> 16#0000;
(* Rosca 1 - horizontal *)
IF bComOK THEN
    r1Anim := s152;
ELSE
    r1Anim := 4;
END_IF;
r1Def := bComOK AND ((w81 AND 16#0020) <> 16#0000);
r1Hor := DWORD_TO_DINT(SHL(WORD_TO_DWORD(INT_TO_WORD(h515)), 16) OR WORD_TO_DWORD(INT_TO_WORD(h514)));
r1Auto := stsAutoRoscas;
r1VelSts := INT_TO_REAL(s151) * 60.0 / 100.0;   (* Hz; UCT em % *)
r1FbLiga := (img013 AND 16#0001) <> 16#0000;
r1FbInt := (img013 AND 16#0020) <> 16#0000;
r1FbRev := (img013 AND 16#0008) <> 16#0000;
(* Rosca 2 - inclinada *)
IF bComOK THEN
    r2Anim := s162;
ELSE
    r2Anim := 4;
END_IF;
r2Def := bComOK AND ((w81 AND 16#0040) <> 16#0000);
r2Hor := DWORD_TO_DINT(SHL(WORD_TO_DWORD(INT_TO_WORD(h517)), 16) OR WORD_TO_DWORD(INT_TO_WORD(h516)));
r2Auto := stsAutoRoscas;
r2VelSts := INT_TO_REAL(s161) * 60.0 / 100.0;   (* Hz; UCT em % *)
r2FbLiga := (img014 AND 16#0001) <> 16#0000;
r2FbInt := (img014 AND 16#0020) <> 16#0000;
r2FbRev := (img014 AND 16#0008) <> 16#0000;

(* ---- 4. Comandos da IHM: troca so o bit comandado na imagem e escreve a palavra ---- *)
IF REQ_PEN_LIGA THEN
    IF penLiga THEN
        img006 := img006 OR 16#0001;
    ELSE
        img006 := img006 AND 16#FFFE;
    END_IF;
    ww006 := WORD_TO_INT(img006);
    CNF_W006 := TRUE;
END_IF;
IF REQ_PEN_INT THEN
    IF penInt THEN
        img006 := img006 OR 16#0020;
    ELSE
        img006 := img006 AND 16#FFDF;
    END_IF;
    ww006 := WORD_TO_INT(img006);
    CNF_W006 := TRUE;
END_IF;
IF REQ_PEN_VEL THEN
    ww101 := REAL_TO_INT(LIMIT(0.0, penVel, 60.0) * 100.0 / 60.0);
    CNF_V101 := TRUE;
END_IF;
IF REQ_B1_LIGA THEN
    IF b1Liga THEN
        img007 := img007 OR 16#0001;
    ELSE
        img007 := img007 AND 16#FFFE;
    END_IF;
    ww007 := WORD_TO_INT(img007);
    CNF_W007 := TRUE;
END_IF;
IF REQ_B1_VEL THEN
    ww116 := REAL_TO_INT(LIMIT(0.0, b1Vel, 60.0) * 100.0 / 60.0);
    CNF_V116 := TRUE;
END_IF;
IF REQ_B2_LIGA THEN
    IF b2Liga THEN
        img008 := img008 OR 16#0001;
    ELSE
        img008 := img008 AND 16#FFFE;
    END_IF;
    ww008 := WORD_TO_INT(img008);
    CNF_W008 := TRUE;
END_IF;
IF REQ_B2_VEL THEN
    ww121 := REAL_TO_INT(LIMIT(0.0, b2Vel, 60.0) * 100.0 / 60.0);
    CNF_V121 := TRUE;
END_IF;
IF REQ_V1_LIGA THEN
    IF v1Liga THEN
        img009 := img009 OR 16#0001;
    ELSE
        img009 := img009 AND 16#FFFE;
    END_IF;
    ww009 := WORD_TO_INT(img009);
    CNF_W009 := TRUE;
END_IF;
IF REQ_V2_LIGA THEN
    IF v2Liga THEN
        img010 := img010 OR 16#0001;
    ELSE
        img010 := img010 AND 16#FFFE;
    END_IF;
    ww010 := WORD_TO_INT(img010);
    CNF_W010 := TRUE;
END_IF;
IF REQ_CMP_LIGA THEN
    IF cmpLiga THEN
        img011 := img011 OR 16#0001;
    ELSE
        img011 := img011 AND 16#FFFE;
    END_IF;
    ww011 := WORD_TO_INT(img011);
    CNF_W011 := TRUE;
END_IF;
IF REQ_CMP_VEL THEN
    ww136 := REAL_TO_INT(LIMIT(0.0, cmpVel, 60.0) * 100.0 / 60.0);
    CNF_V136 := TRUE;
END_IF;
IF REQ_RSP_LIGA THEN
    IF rspLiga THEN
        img012 := img012 OR 16#0001;
    ELSE
        img012 := img012 AND 16#FFFE;
    END_IF;
    ww012 := WORD_TO_INT(img012);
    CNF_W012 := TRUE;
END_IF;
IF REQ_RSP_INT THEN
    IF rspInt THEN
        img012 := img012 OR 16#0020;
    ELSE
        img012 := img012 AND 16#FFDF;
    END_IF;
    ww012 := WORD_TO_INT(img012);
    CNF_W012 := TRUE;
END_IF;
IF REQ_RSP_REV THEN
    IF rspRev THEN
        img012 := img012 OR 16#0008;
    ELSE
        img012 := img012 AND 16#FFF7;
    END_IF;
    ww012 := WORD_TO_INT(img012);
    CNF_W012 := TRUE;
END_IF;
IF REQ_RSP_VEL THEN
    ww141 := REAL_TO_INT(LIMIT(0.0, rspVel, 60.0) * 100.0 / 60.0);
    CNF_V141 := TRUE;
END_IF;
IF REQ_R1_LIGA THEN
    IF r1Liga THEN
        img013 := img013 OR 16#0001;
    ELSE
        img013 := img013 AND 16#FFFE;
    END_IF;
    ww013 := WORD_TO_INT(img013);
    CNF_W013 := TRUE;
END_IF;
IF REQ_R1_INT THEN
    IF r1Int THEN
        img013 := img013 OR 16#0020;
    ELSE
        img013 := img013 AND 16#FFDF;
    END_IF;
    ww013 := WORD_TO_INT(img013);
    CNF_W013 := TRUE;
END_IF;
IF REQ_R1_REV THEN
    IF r1Rev THEN
        img013 := img013 OR 16#0008;
    ELSE
        img013 := img013 AND 16#FFF7;
    END_IF;
    ww013 := WORD_TO_INT(img013);
    CNF_W013 := TRUE;
END_IF;
IF REQ_R1_VEL THEN
    ww151 := REAL_TO_INT(LIMIT(0.0, r1Vel, 60.0) * 100.0 / 60.0);
    CNF_V151 := TRUE;
END_IF;
IF REQ_R2_LIGA THEN
    IF r2Liga THEN
        img014 := img014 OR 16#0001;
    ELSE
        img014 := img014 AND 16#FFFE;
    END_IF;
    ww014 := WORD_TO_INT(img014);
    CNF_W014 := TRUE;
END_IF;
IF REQ_R2_INT THEN
    IF r2Int THEN
        img014 := img014 OR 16#0020;
    ELSE
        img014 := img014 AND 16#FFDF;
    END_IF;
    ww014 := WORD_TO_INT(img014);
    CNF_W014 := TRUE;
END_IF;
IF REQ_R2_REV THEN
    IF r2Rev THEN
        img014 := img014 OR 16#0008;
    ELSE
        img014 := img014 AND 16#FFF7;
    END_IF;
    ww014 := WORD_TO_INT(img014);
    CNF_W014 := TRUE;
END_IF;
IF REQ_R2_VEL THEN
    ww161 := REAL_TO_INT(LIMIT(0.0, r2Vel, 60.0) * 100.0 / 60.0);
    CNF_V161 := TRUE;
END_IF;
IF REQ_LIGA_PEN THEN
    IF hmiLigaPeneira THEN
        img015 := img015 OR 16#0001;
    ELSE
        img015 := img015 AND 16#FFFE;
    END_IF;
    ww015 := WORD_TO_INT(img015);
    CNF_W015 := TRUE;
END_IF;
IF REQ_SEL_PEN THEN
    IF hmiSelPeneira THEN
        img015 := img015 OR 16#0004;
    ELSE
        img015 := img015 AND 16#FFFB;
    END_IF;
    ww015 := WORD_TO_INT(img015);
    CNF_W015 := TRUE;
END_IF;
IF REQ_LIGA_ROS THEN
    IF hmiLigaRoscas THEN
        img016 := img016 OR 16#0001;
    ELSE
        img016 := img016 AND 16#FFFE;
    END_IF;
    ww016 := WORD_TO_INT(img016);
    CNF_W016 := TRUE;
END_IF;
IF REQ_SEL_ROS THEN
    IF hmiSelRoscas THEN
        img016 := img016 OR 16#0004;
    ELSE
        img016 := img016 AND 16#FFFB;
    END_IF;
    ww016 := WORD_TO_INT(img016);
    CNF_W016 := TRUE;
END_IF;
IF REQ_LIGA_RC THEN
    IF hmiLigaRaspComp THEN
        img017 := img017 OR 16#0001;
    ELSE
        img017 := img017 AND 16#FFFE;
    END_IF;
    ww017 := WORD_TO_INT(img017);
    CNF_W017 := TRUE;
END_IF;
IF REQ_SEL_RC THEN
    IF hmiSelRaspComp THEN
        img017 := img017 OR 16#0004;
    ELSE
        img017 := img017 AND 16#FFFB;
    END_IF;
    ww017 := WORD_TO_INT(img017);
    CNF_W017 := TRUE;
END_IF;
IF REQ_SEL_BOMBA THEN
    IF hmiSelBomba THEN
        img007 := img007 OR 16#0008;
    ELSE
        img007 := img007 AND 16#FFF7;
    END_IF;
    ww007 := WORD_TO_INT(img007);
    CNF_W007 := TRUE;
END_IF;

(* ---- 5. Reset: pulso em 40005.3, bomba de gordura e reconhecimento ---- *)
bReset := (REQ_RESET AND hmiReset) OR (REQ_RESET_PROC AND cmdResetFalhas);
IF bReset THEN
    img005 := img005 OR 16#0008;
    ww005 := WORD_TO_INT(img005);
    CNF_W005 := TRUE;
    uSegReset := cfgTempoReset;
    IF uSegReset = 0 THEN
        uSegReset := 1;
    END_IF;
    resetBomba := TRUE;
    CNF_RESET := TRUE;
ELSIF TICK AND uSegReset > 0 THEN
    uSegReset := uSegReset - 1;
    IF uSegReset = 0 THEN
        img005 := img005 AND 16#FFF7;
        ww005 := WORD_TO_INT(img005);
        CNF_W005 := TRUE;
    END_IF;
END_IF;

(* ---- 6. Disponibilidade (condicoes para o AND editavel do CAT) e cadeia das UCTs ---- *)
habilitada := cfgInstalada AND stpHabilitada;
okComunicacao := bComOK;
okEmergencia := bComOK AND NOT stsEmergenciaUCT;
okPeneira := bComOK AND NOT penDef;
okMotores := bComOK AND NOT (b1Def OR b2Def OR cmpDef OR rspDef OR r1Def OR r2Def);
stsDisponivel := disponivel AND habilitada;
stsAlgumaHabilitada := habilitada OR antHabilitada;
stsAlgumaDisponivel := stsDisponivel OR antDisponivel;
stsBloqueioEEE := stsAlgumaHabilitada AND NOT stsAlgumaDisponivel;

(* ---- 7. Bomba de gordura e valvula de lavagem ---- *)
bNivelAltoG := stsNivelAltoGordura;
IF emergencia OR NOT bombaAutomatico THEN
    uEtapa := 0;
    uSegEtapa := 0;
    uSegValv := 0;
    cmdLigarBomba := FALSE;
    bValvAuto := FALSE;
ELSE
    IF TICK THEN
        uSegEtapa := uSegEtapa + 1;
        IF uEtapa >= 2 THEN
            uSegValv := uSegValv + 1;
        END_IF;
    END_IF;
    IF uEtapa = 0 THEN
        IF bNivelAltoG THEN
            uEtapa := 1;
            uSegEtapa := 0;
        END_IF;
    END_IF;
    IF uEtapa = 1 THEN
        IF uSegEtapa >= UINT_TO_UDINT(stpTempoPreLavagem) THEN
            uEtapa := 2;
            uSegEtapa := 0;
            uSegValv := 0;
        END_IF;
    END_IF;
    IF uEtapa = 2 THEN
        IF NOT bNivelAltoG THEN
            uEtapa := 3;
            uSegEtapa := 0;
        END_IF;
    ELSIF uEtapa = 3 THEN
        IF bNivelAltoG THEN
            uEtapa := 2;
            uSegEtapa := 0;
        ELSIF uSegEtapa >= UINT_TO_UDINT(stpTempoDesliga) THEN
            uEtapa := 0;
            uSegEtapa := 0;
        END_IF;
    END_IF;
    cmdLigarBomba := uEtapa >= 2;
    bValvAuto := (uEtapa = 1) OR (uEtapa >= 2 AND uSegValv < UINT_TO_UDINT(stpTempoValvula));
END_IF;
stpVelBombaOut := stpVelBomba / 0.6;   (* IHM/SCADA em Hz -> % do Motor_Generico *)
IF emergencia THEN
    cmdValvula := FALSE;
ELSIF bombaAutomatico THEN
    cmdValvula := bValvAuto;
ELSE
    cmdValvula := hmiValvula;
END_IF;
stsValvula := cmdValvula;
IF NOT bombaAutomatico THEN
    stsEtapaGordura := 4;
ELSE
    stsEtapaGordura := uEtapa;
END_IF;
IF bombaAutomatico AND uEtapa = 1 THEN
    stsTempoRestante := UDINT_TO_INT(UINT_TO_UDINT(stpTempoPreLavagem) - MIN(uSegEtapa, UINT_TO_UDINT(stpTempoPreLavagem)));
ELSIF bombaAutomatico AND uEtapa = 3 THEN
    stsTempoRestante := UDINT_TO_INT(UINT_TO_UDINT(stpTempoDesliga) - MIN(uSegEtapa, UINT_TO_UDINT(stpTempoDesliga)));
ELSE
    stsTempoRestante := 0;
END_IF;

(* ---- 8. Alarmes (UCT nao instalada nao alarma) ---- *)
almCom := stsFalhaComunicacao;
almEmergencia := stsEmergenciaUCT;
almDefPEN := penDef;
almDefB1 := b1Def;
almDefB2 := b2Def;
almDefCMP := cmpDef;
almDefRSP := rspDef;
almDefR1 := r1Def;
almDefR2 := r2Def;
almNivelAgua := stsNivelBaixoAgua;
almNivelPeneira := stsNivelAltoPeneira;
stsAlarme := almCom OR almEmergencia OR almDefPEN OR almDefB1 OR almDefB2 OR almDefCMP OR almDefRSP OR almDefR1 OR almDefR2 OR almNivelAgua OR almNivelPeneira;

(* ---- 9. Eventos so na mudanca ---- *)
wD := 0;
IF okEmergencia THEN wD := wD OR 16#0001; END_IF;
IF okPeneira THEN wD := wD OR 16#0002; END_IF;
IF okMotores THEN wD := wD OR 16#0004; END_IF;
IF okComunicacao THEN wD := wD OR 16#0008; END_IF;
IF habilitada THEN wD := wD OR 16#0010; END_IF;
CNF_DISP := initPass OR (wD <> oldD);
wP := 0;
IF stsDisponivel THEN wP := wP OR 16#00000001; END_IF;
IF stsAlgumaHabilitada THEN wP := wP OR 16#00000002; END_IF;
IF stsAlgumaDisponivel THEN wP := wP OR 16#00000004; END_IF;
IF stsBloqueioEEE THEN wP := wP OR 16#00000008; END_IF;
IF stsFalhaComunicacao THEN wP := wP OR 16#00000010; END_IF;
IF stsEmergenciaUCT THEN wP := wP OR 16#00000020; END_IF;
IF stsNivelAltoGordura THEN wP := wP OR 16#00000040; END_IF;
IF stsAlarme THEN wP := wP OR 16#00000080; END_IF;
IF stsNivelBaixoPeneira THEN wP := wP OR 16#00000100; END_IF;
IF stsNivelAltoPeneira THEN wP := wP OR 16#00000200; END_IF;
IF stsNivelBaixoAgua THEN wP := wP OR 16#00000400; END_IF;
IF stsAutoPeneira THEN wP := wP OR 16#00000800; END_IF;
IF stsAutoRoscas THEN wP := wP OR 16#00001000; END_IF;
IF stsAutoRaspComp THEN wP := wP OR 16#00002000; END_IF;
IF stsLigaAutoPeneira THEN wP := wP OR 16#00004000; END_IF;
IF stsLigaAutoRoscas THEN wP := wP OR 16#00008000; END_IF;
IF stsLigaAutoRaspComp THEN wP := wP OR 16#00010000; END_IF;
IF stsSelecaoBomba THEN wP := wP OR 16#00020000; END_IF;
IF stsValvula THEN wP := wP OR 16#00040000; END_IF;
CNF := initPass OR ((wP AND 16#000000FF) <> (oldP AND 16#000000FF));
bMudou := (wP <> oldP) OR (wD <> oldD);
oldD := wD;                                (* depois do bMudou: mudanca so em wD tambem atualiza a IHM *)
IF stsNivelPeneira <> o_stsNivelPeneira THEN bMudou := TRUE; o_stsNivelPeneira := stsNivelPeneira; END_IF;
IF stsEtapaGordura <> o_stsEtapaGordura THEN bMudou := TRUE; o_stsEtapaGordura := stsEtapaGordura; END_IF;
IF stsTempoRestante <> o_stsTempoRestante THEN bMudou := TRUE; o_stsTempoRestante := stsTempoRestante; END_IF;
CNF_HMI := initPass OR bMudou;
oldP := wP;
bMudou := FALSE;
IF penAnim <> o_penAnim THEN bMudou := TRUE; o_penAnim := penAnim; END_IF;
IF penDef <> o_penDef THEN bMudou := TRUE; o_penDef := penDef; END_IF;
IF penHor <> o_penHor THEN bMudou := TRUE; o_penHor := penHor; END_IF;
IF penAuto <> o_penAuto THEN bMudou := TRUE; o_penAuto := penAuto; END_IF;
IF penVelSts <> o_penVelSts THEN bMudou := TRUE; o_penVelSts := penVelSts; END_IF;
IF penFbLiga <> o_penFbLiga THEN bMudou := TRUE; o_penFbLiga := penFbLiga; END_IF;
IF penFbInt <> o_penFbInt THEN bMudou := TRUE; o_penFbInt := penFbInt; END_IF;
IF penFbRev <> o_penFbRev THEN bMudou := TRUE; o_penFbRev := penFbRev; END_IF;
IF b1Anim <> o_b1Anim THEN bMudou := TRUE; o_b1Anim := b1Anim; END_IF;
IF b1Def <> o_b1Def THEN bMudou := TRUE; o_b1Def := b1Def; END_IF;
IF b1Hor <> o_b1Hor THEN bMudou := TRUE; o_b1Hor := b1Hor; END_IF;
IF b1Auto <> o_b1Auto THEN bMudou := TRUE; o_b1Auto := b1Auto; END_IF;
IF b1VelSts <> o_b1VelSts THEN bMudou := TRUE; o_b1VelSts := b1VelSts; END_IF;
IF b1FbLiga <> o_b1FbLiga THEN bMudou := TRUE; o_b1FbLiga := b1FbLiga; END_IF;
IF b1FbInt <> o_b1FbInt THEN bMudou := TRUE; o_b1FbInt := b1FbInt; END_IF;
IF b1FbRev <> o_b1FbRev THEN bMudou := TRUE; o_b1FbRev := b1FbRev; END_IF;
IF b2Anim <> o_b2Anim THEN bMudou := TRUE; o_b2Anim := b2Anim; END_IF;
IF b2Def <> o_b2Def THEN bMudou := TRUE; o_b2Def := b2Def; END_IF;
IF b2Hor <> o_b2Hor THEN bMudou := TRUE; o_b2Hor := b2Hor; END_IF;
IF b2Auto <> o_b2Auto THEN bMudou := TRUE; o_b2Auto := b2Auto; END_IF;
IF b2VelSts <> o_b2VelSts THEN bMudou := TRUE; o_b2VelSts := b2VelSts; END_IF;
IF b2FbLiga <> o_b2FbLiga THEN bMudou := TRUE; o_b2FbLiga := b2FbLiga; END_IF;
IF b2FbInt <> o_b2FbInt THEN bMudou := TRUE; o_b2FbInt := b2FbInt; END_IF;
IF b2FbRev <> o_b2FbRev THEN bMudou := TRUE; o_b2FbRev := b2FbRev; END_IF;
IF v1Anim <> o_v1Anim THEN bMudou := TRUE; o_v1Anim := v1Anim; END_IF;
IF v1Def <> o_v1Def THEN bMudou := TRUE; o_v1Def := v1Def; END_IF;
IF v1Hor <> o_v1Hor THEN bMudou := TRUE; o_v1Hor := v1Hor; END_IF;
IF v1Auto <> o_v1Auto THEN bMudou := TRUE; o_v1Auto := v1Auto; END_IF;
IF v1VelSts <> o_v1VelSts THEN bMudou := TRUE; o_v1VelSts := v1VelSts; END_IF;
IF v1FbLiga <> o_v1FbLiga THEN bMudou := TRUE; o_v1FbLiga := v1FbLiga; END_IF;
IF v1FbInt <> o_v1FbInt THEN bMudou := TRUE; o_v1FbInt := v1FbInt; END_IF;
IF v1FbRev <> o_v1FbRev THEN bMudou := TRUE; o_v1FbRev := v1FbRev; END_IF;
IF v2Anim <> o_v2Anim THEN bMudou := TRUE; o_v2Anim := v2Anim; END_IF;
IF v2Def <> o_v2Def THEN bMudou := TRUE; o_v2Def := v2Def; END_IF;
IF v2Hor <> o_v2Hor THEN bMudou := TRUE; o_v2Hor := v2Hor; END_IF;
IF v2Auto <> o_v2Auto THEN bMudou := TRUE; o_v2Auto := v2Auto; END_IF;
IF v2VelSts <> o_v2VelSts THEN bMudou := TRUE; o_v2VelSts := v2VelSts; END_IF;
IF v2FbLiga <> o_v2FbLiga THEN bMudou := TRUE; o_v2FbLiga := v2FbLiga; END_IF;
IF v2FbInt <> o_v2FbInt THEN bMudou := TRUE; o_v2FbInt := v2FbInt; END_IF;
IF v2FbRev <> o_v2FbRev THEN bMudou := TRUE; o_v2FbRev := v2FbRev; END_IF;
IF cmpAnim <> o_cmpAnim THEN bMudou := TRUE; o_cmpAnim := cmpAnim; END_IF;
IF cmpDef <> o_cmpDef THEN bMudou := TRUE; o_cmpDef := cmpDef; END_IF;
IF cmpHor <> o_cmpHor THEN bMudou := TRUE; o_cmpHor := cmpHor; END_IF;
IF cmpAuto <> o_cmpAuto THEN bMudou := TRUE; o_cmpAuto := cmpAuto; END_IF;
IF cmpVelSts <> o_cmpVelSts THEN bMudou := TRUE; o_cmpVelSts := cmpVelSts; END_IF;
IF cmpFbLiga <> o_cmpFbLiga THEN bMudou := TRUE; o_cmpFbLiga := cmpFbLiga; END_IF;
IF cmpFbInt <> o_cmpFbInt THEN bMudou := TRUE; o_cmpFbInt := cmpFbInt; END_IF;
IF cmpFbRev <> o_cmpFbRev THEN bMudou := TRUE; o_cmpFbRev := cmpFbRev; END_IF;
IF rspAnim <> o_rspAnim THEN bMudou := TRUE; o_rspAnim := rspAnim; END_IF;
IF rspDef <> o_rspDef THEN bMudou := TRUE; o_rspDef := rspDef; END_IF;
IF rspHor <> o_rspHor THEN bMudou := TRUE; o_rspHor := rspHor; END_IF;
IF rspAuto <> o_rspAuto THEN bMudou := TRUE; o_rspAuto := rspAuto; END_IF;
IF rspVelSts <> o_rspVelSts THEN bMudou := TRUE; o_rspVelSts := rspVelSts; END_IF;
IF rspFbLiga <> o_rspFbLiga THEN bMudou := TRUE; o_rspFbLiga := rspFbLiga; END_IF;
IF rspFbInt <> o_rspFbInt THEN bMudou := TRUE; o_rspFbInt := rspFbInt; END_IF;
IF rspFbRev <> o_rspFbRev THEN bMudou := TRUE; o_rspFbRev := rspFbRev; END_IF;
IF r1Anim <> o_r1Anim THEN bMudou := TRUE; o_r1Anim := r1Anim; END_IF;
IF r1Def <> o_r1Def THEN bMudou := TRUE; o_r1Def := r1Def; END_IF;
IF r1Hor <> o_r1Hor THEN bMudou := TRUE; o_r1Hor := r1Hor; END_IF;
IF r1Auto <> o_r1Auto THEN bMudou := TRUE; o_r1Auto := r1Auto; END_IF;
IF r1VelSts <> o_r1VelSts THEN bMudou := TRUE; o_r1VelSts := r1VelSts; END_IF;
IF r1FbLiga <> o_r1FbLiga THEN bMudou := TRUE; o_r1FbLiga := r1FbLiga; END_IF;
IF r1FbInt <> o_r1FbInt THEN bMudou := TRUE; o_r1FbInt := r1FbInt; END_IF;
IF r1FbRev <> o_r1FbRev THEN bMudou := TRUE; o_r1FbRev := r1FbRev; END_IF;
IF r2Anim <> o_r2Anim THEN bMudou := TRUE; o_r2Anim := r2Anim; END_IF;
IF r2Def <> o_r2Def THEN bMudou := TRUE; o_r2Def := r2Def; END_IF;
IF r2Hor <> o_r2Hor THEN bMudou := TRUE; o_r2Hor := r2Hor; END_IF;
IF r2Auto <> o_r2Auto THEN bMudou := TRUE; o_r2Auto := r2Auto; END_IF;
IF r2VelSts <> o_r2VelSts THEN bMudou := TRUE; o_r2VelSts := r2VelSts; END_IF;
IF r2FbLiga <> o_r2FbLiga THEN bMudou := TRUE; o_r2FbLiga := r2FbLiga; END_IF;
IF r2FbInt <> o_r2FbInt THEN bMudou := TRUE; o_r2FbInt := r2FbInt; END_IF;
IF r2FbRev <> o_r2FbRev THEN bMudou := TRUE; o_r2FbRev := r2FbRev; END_IF;
CNF_EQ := initPass OR bMudou;
wA := 0;
IF almCom THEN wA := wA OR 16#0001; END_IF;
IF almEmergencia THEN wA := wA OR 16#0002; END_IF;
IF almDefPEN THEN wA := wA OR 16#0004; END_IF;
IF almDefB1 THEN wA := wA OR 16#0008; END_IF;
IF almDefB2 THEN wA := wA OR 16#0010; END_IF;
IF almDefCMP THEN wA := wA OR 16#0020; END_IF;
IF almDefRSP THEN wA := wA OR 16#0040; END_IF;
IF almDefR1 THEN wA := wA OR 16#0080; END_IF;
IF almDefR2 THEN wA := wA OR 16#0100; END_IF;
IF almNivelAgua THEN wA := wA OR 16#0200; END_IF;
IF almNivelPeneira THEN wA := wA OR 16#0400; END_IF;
CNF_ALM := initPass OR (wA <> oldA);
oldA := wA;
CNF_BOMBA := initPass OR (cmdLigarBomba <> oldLigB) OR (stpVelBombaOut <> oldVelB);
oldLigB := cmdLigarBomba;
oldVelB := stpVelBombaOut;
CNF_VALVULA := initPass OR (cmdValvula <> oldValv);
oldValv := cmdValvula;
initPass := FALSE;
  END_ALGORITHM
END_FUNCTION_BLOCK
